    rq_activate_all_grippers(False)
    # end: URCap Program Node
  else:
    $ 55 "Else" "noBreak"
    # begin: URCap Program Node
    #   Source: Robotiq_Grippers, 3.17.0.105337, Robotiq Inc.
    #   Type: Gripper Activate
    $ 56 "Gripper Reset and Activate"

    kill rq_gripper_communication_thread
    rq_gripper_communication_thread_started = False
    rq_close_gripper_socket("1")
    rq_close_gripper_socket("2")
    rq_close_gripper_socket("3")
    rq_close_gripper_socket("4")

    rq_init_comm_if_connected(9, "1")
    rq_init_comm_if_connected(2, "2")
    rq_init_comm_if_connected(3, "3")
    rq_init_comm_if_connected(4, "4")
    rq_print_connected_grippers()
    rq_gripper_communication_thread = run rq_gripper_communication()

    while(not rq_gripper_communication_thread_started):
        sleep(0.008)
    end

    rq_set_max_current_for_all_grippers()

    reset_and_activate = True

    rq_activate_all_grippers(True)
    # end: URCap Program Node
  end
  $ 57 "zero_ftsensor()"
  zero_ftsensor()
  $ 58 "EXTT"
  $ 59 "Set GRP_3F_Enable=Off"
  set_standard_digital_out(4, False)
  $ 60 "Set BarcodeTrigger=Off"
  set_standard_digital_out(6, False)
  $ 61 "Set GRP_3F_Decap=Off"
  set_standard_digital_out(3, False)
  $ 62 "Set GRP_3F_Cap=Off"
  set_standard_digital_out(2, False)
  $ 63 "Set GRP_3F_Open=Off"
  set_standard_digital_out(5, False)
  $ 64 "PSE_T≔get_tool_free_pose(dir=[0,0,0.150], move_in_base_frame=True)"
  global PSE_T=get_tool_free_pose(dir=[0,0,0.150], move_in_base_frame=True)
  $ 65 "If is_reachable(Base_const, [PSE_T])"
  if (is_reachable(p[0.0,0.0,0.0,0.0,0.0,0.0], [PSE_T])):
    $ 66 "MoveL"
    $ 67 "PSE_T" "breakAfter"
    movel(PSE_T, a=1.2, v=0.15)
  end
  $ 68 "powder dispensing variable init"
  $ 69 "Start_thread≔ False "
  global Start_thread=  False
  $ 70 "vib_thread≔ False "
  global vib_thread=  False
  $ 71 "w_full_thread≔ False "
  global w_full_thread=  False
  $ 72 "d_cc≔0.07"
  global d_cc=0.07
  $ 73 "kp≔0.0035"
  global kp=0.0035
  $ 74 "ki≔0.0001"
  global ki=0.0001
  $ 75 "kd≔0.003"
  global kd=0.003
  $ 76 "dt≔0.2"
  global dt=0.2
  $ 77 "Integral_error≔0"
  global Integral_error=0
  $ 78 "current_error≔0"
  global current_error=0
  $ 79 "previous_error≔0"
  global previous_error=0
  $ 80 "tilt_increment≔0"
  global tilt_increment=0
  $ 81 "tilt_angle≔0"
  global tilt_angle=0
  $ 82 "diff≔0"
  global diff=0
  $ 83 "tilt_to_home()"
  tilt_to_home()
  $ 84 "tilt_to_home()"
  tilt_to_home()
  $ 85 "switch_spat_M≔ True "
  global switch_spat_M=  True
  $ 86 "switch_spat_S≔ True "
  global switch_spat_S=  True
  $ 87 "switch_spat_F_M≔ True "
  global switch_spat_F_M=  True
  $ 88 "switch_spat_F_S≔ True "
  global switch_spat_F_S=  True
  $ 89 "last_scale≔0"
  global last_scale=0
  $ 818 "Thread_1"
  thread Thread_1():
    while (True):
      $ 819 "Dosing Weight"
      $ 820 "If Start_thread≟ True "
      if (Start_thread ==   True  ):
        $ 821 "weight_value≔get_weight()"
        global weight_value=get_weight()
        $ 822 "diff≔target_weight-weight_value"
        global diff=target_weight-weight_value
        $ 823 "Wait: 0.2"
        sleep(0.2)
        $ 824 "sync()"
        sync()
      end
      $ 825 "sync()"
      sync()
    end
  end
  threadId_Thread_1 = run Thread_1()
  $ 826 "Thread_2"
  thread Thread_2():
    while (True):
      $ 827 "Vibration motor"
      $ 828 "Loop vib_thread≟ True "
      thread Thread_while_828():
        while (True):
          $ 829 "diff≔target_weight-weight_value"
          global diff=target_weight-weight_value
          $ 830 "If diff>0.02 and spatula≠'spatula_flat_S' "
          global thread_flag_830=0
          thread Thread_if_830():
            $ 832 "Set AO[0]=4.0"
            set_standard_analog_out(0, 0.4)
            thread_flag_830 = 1
          end
          if (diff>0.02  and  spatula != "spatula_flat_S" ):
            global thread_handler_830=run Thread_if_830()
            while (thread_flag_830 == 0):
              if not(diff>0.02  and  spatula != "spatula_flat_S" ):
                kill thread_handler_830
                thread_flag_830 = 2
              else:
                sync()
              end
            end
          else:
            thread_flag_830 = 2
          end
          if (thread_flag_830 == 2):
            $ 833 "ElseIf diff>0.02 and spatula≟'spatula_flat_S'"
            if (diff>0.02 and spatula == "spatula_flat_S"):
              $ 834 "vibration_3()"
              vibration_3()
            else:
              $ 835 "ElseIf diff≤0.03"
              global thread_flag_835=0
              thread Thread_if_835():
                $ 836 "vibration_2()"
                vibration_2()
                thread_flag_835 = 1
              end
              if (diff <= 0.03):
                global thread_handler_835=run Thread_if_835()
                while (thread_flag_835 == 0):
                  if not(diff <= 0.03):
                    kill thread_handler_835
                    thread_flag_835 = 2
                  else:
                    sync()
                  end
                end
              else:
                thread_flag_835 = 2
              end
              if (thread_flag_835 == 2):
                $ 837 "Else" "noBreak"
                $ 838 "Set AO[0]=0.0"
                set_standard_analog_out(0, 0.0)
              end
            end
          end
        end
      end
      if (vib_thread ==   True  ):
        global thread_handler_828=run Thread_while_828()
        while (vib_thread ==   True  ):
          sync()
        end
        kill thread_handler_828
      end
      $ 839 "sync()"
      sync()
    end
  end
  threadId_Thread_2 = run Thread_2()
  $ 840 "Thread_3"
  thread Thread_3():
    while (True):
      $ 841 "Container weight"
      $ 842 "If w_full_thread≟ True "
      if (w_full_thread ==   True  ):
        $ 843 "aa_weight_cont≔get_cont_weight()"
        global aa_weight_cont=get_cont_weight()
        $ 844 "Wait: 0.2"
        sleep(0.2)
        $ 845 "sync()"
        sync()
      end
      $ 846 "sync()"
      sync()
    end
  end
  threadId_Thread_3 = run Thread_3()
  while (True):
    $ 90 "Robot Program"
    $ 91 "MAIN"
    $ 92 "command_manager(external_control='uGO', cond_suspend=(ITM_Manipulated and AMR_AtTarget and AMR_Charging and AMR_Battery<40), cond_unsuspend=(AMR_Battery≟60))"
    command_manager(external_control="uGO", cond_suspend=(ITM_Manipulated  and  AMR_AtTarget  and  AMR_Charging  and  AMR_Battery<40), cond_unsuspend=(AMR_Battery == 60))
    $ 93 "log_state(STATE_Info)"
    log_state(STATE_Info)
    $ 94 "Switch STATE"
    switch_1 = STATE
    $ 95 "Case 1"
    if (1 == switch_1):
      $ 96 "Stopping"
      $ 97 "STATE_Info≔'Stopping'"
      global STATE_Info="Stopping"
      $ 98 "end_freedrive_mode()"
      end_freedrive_mode()
      $ 99 "Set"
      set_tcp(p[0.0,0.0,0.161,3.1415,0.0,0.0])
      $ 100 "PSE_T≔get_tool_free_pose(dir=[0,0,0.150], move_in_base_frame=True)"
      global PSE_T=get_tool_free_pose(dir=[0,0,0.150], move_in_base_frame=True)
      $ 101 "If is_reachable(Base_const, [PSE_T])"
      if (is_reachable(p[0.0,0.0,0.0,0.0,0.0,0.0], [PSE_T])):
        $ 102 "MoveL"
        $ 103 "PSE_T" "breakAfter"
        movel(PSE_T, a=1.2, v=0.15)
      end
      $ 104 "do_transition(keep_rxry=OBJ_Picked, r=0)"
      do_transition(keep_rxry=OBJ_Picked, r=0)
      $ 113 "Call Sub_AMR_MiR_V3"
      Sub_AMR_MiR_V3()
      $ 114 "If stopping() and AMR_Done"
      if (stopping()  and  AMR_Done):
        $ 115 "STATE≔2"
        global STATE=2
        $ 116 "ugo_update_outputs()"
        ugo_update_outputs()
      end
    elif (2 == switch_1):
      $ 117 "Case 2"
      $ 118 "Stopped"
      $ 119 "STATE_Info≔'Stopped'"
      global STATE_Info="Stopped"
      $ 120 "Call Sub_AMR_MiR_V3"
      Sub_AMR_MiR_V3()
      $ 121 "If CMD_Reset  or PB_Start"
      if (CMD_Reset   or  get_standard_digital_in(0)):
        $ 122 "STATE≔3"
        global STATE=3
        $ 123 "ugo_update_outputs()"
        ugo_update_outputs()
      end
    elif (3 == switch_1):
      $ 124 "Case 3"
      $ 125 " Resetting"
      $ 126 "STATE_Info≔'Resetting'"
      global STATE_Info="Resetting"
      $ 127 "uML"
      $ 128 "reset_error()"
      reset_error()
      $ 129 "reset_warning()"
      reset_warning()
      $ 130 "PROCESS_Step≔0"
      global PROCESS_Step=0
      $ 131 "PROCESS_Info≔''"
      global PROCESS_Info=""
      $ 132 "ARM_Referenced≔ False "
      global ARM_Referenced=  False
      $ 133 "WRK_Done≔ False "
      global WRK_Done=  False
      $ 134 "ITM_Prepared≔ False "
      global ITM_Prepared=  False
      $ 135 "ITM_Manipulated≔ False "
      global ITM_Manipulated=  False
      $ 136 "STP≔0"
      global STP=0
      $ 137 "Action≔0"
      global Action=0
      $ 138 "Action_Info≔''"
      global Action_Info=""
      $ 139 "ITM_ID≔0"
      global ITM_ID=0
      $ 140 "JIG≔0"
      global JIG=0
      $ 141 "JIG_Slot≔0"
      global JIG_Slot=0
      $ 142 "Task_info≔''"
      global Task_info=""
      $ 143 "Set"
      set_tcp(p[0.0,0.0,0.161,3.1415,0.0,0.0])
      $ 144 "App"
      $ 145 "'ADD APPLICATION SPECIFIC COMMANDS'"
      # 'ADD APPLICATION SPECIFIC COMMANDS'
      $ 146 "OBJ_Type≔0"
      global OBJ_Type=0
      $ 147 "OBJ_Nbr≔0"
      global OBJ_Nbr=0
      $ 148 "If CNT_Rack_Output≥50"
      if (CNT_Rack_Output >= 50):
        $ 149 "CNT_Rack_Output≔0"
        global CNT_Rack_Output=0
      end
      $ 150 "TASK≔struct(ID=0, NAVI=struct(target=0, footprint=0, protectiveOff=0, dock=0), WORK=struct(ITM_ID_Src=0, JIG_ID_Src=0, OBJ_Nbr_Src=0, ACT_Src=0, ITM_ID_Tgt=0, JIG_ID_Tgt=0, OBJ_Nbr_Tgt=0, ACT_Tgt=0, OBJ_Type=0))"
      global TASK=struct(ID=0, NAVI=struct(target=0, footprint=0, protectiveOff=0, dock=0), WORK=struct(ITM_ID_Src=0, JIG_ID_Src=0, OBJ_Nbr_Src=0, ACT_Src=0, ITM_ID_Tgt=0, JIG_ID_Tgt=0, OBJ_Nbr_Tgt=0, ACT_Tgt=0, OBJ_Type=0))
      $ 151 "Call Sub_AMR_MiR_V3"
      Sub_AMR_MiR_V3()
      $ 152 "If resetting() and AMR_Done"
      if (resetting()  and  AMR_Done):
        $ 153 "STATE≔4"
        global STATE=4
        $ 154 "ugo_update_outputs()"
        ugo_update_outputs()
      end
    elif (4 == switch_1):
      $ 155 "Case 4"
      $ 156 "Idle"
      $ 157 "STATE_Info≔'Idle'"
      global STATE_Info="Idle"
      $ 158 "If CMD_Start"
      if (CMD_Start):
        $ 159 "STATE≔5"
        global STATE=5
        $ 160 "ugo_update_outputs()"
        ugo_update_outputs()
      end
    elif (5 == switch_1):
      $ 161 "Case 5"
      $ 162 "Starting"
      $ 163 "STATE_Info≔'Starting'"
      global STATE_Info="Starting"
      $ 164 "'ADD COMMANDS WHAT TO START WITH'"
      # 'ADD COMMANDS WHAT TO START WITH'
      $ 165 "Call Sub_AMR_MiR_V3"
      Sub_AMR_MiR_V3()
      $ 166 "get ugo data"
      $ 167 "Assign Tasks"
      $ 168 "TASK.ID = ugo_get_task()"
      TASK.ID = ugo_get_task()
      $ 169 "If TASK.ID≟1"
      if (TASK.ID == 1):
        $ 170 "Task_info≔'Charge'"
        global Task_info="Charge"
        $ 171 "Parameters"
        $ 172 "AMR_PosTarget≔1"
        global AMR_PosTarget=1
      else:
        $ 173 "ElseIf TASK.ID≟9"
        if (TASK.ID == 9):
          $ 174 "'Pick Sarstedt Rack from Variable source'"
          # 'Pick Sarstedt Rack from Variable source'
          $ 175 "Task_info≔'Navigate to Target'"
          global Task_info="Navigate to Target"
          $ 176 "Parameters"
          $ 177 "AMR_PosTarget≔UGO.read_input('00','ITM_ID')"
          global AMR_PosTarget=UGO.read_input("00","ITM_ID")
        else:
          $ 178 "ElseIf TASK.ID≟13"
          if (TASK.ID == 13):
            $ 179 "Task_info≔'Dose Powder'"
            global Task_info="Dose Powder"
            $ 180 "Parameters"
            $ 181 "ITM_ID≔1"
            global ITM_ID=1
            $ 182 "W_now≔(UGO.read_input('00','Container_weight'))/1000"
            global W_now=(UGO.read_input("00","Container_weight"))/1000
            $ 183 "Pow_name≔(UGO.read_input('00','Powder_name'))"
            global Pow_name=(UGO.read_input("00","Powder_name"))
            $ 184 "target_weight≔(UGO.read_input('00','Target_weight'))/1000"
            global target_weight=(UGO.read_input("00","Target_weight"))/1000
            $ 185 "send_picking_info(Pow_name,target_weight)"
            send_picking_info(Pow_name,target_weight)
            $ 186 "w_dosed_total≔0"
            global w_dosed_total=0
            $ 187 "OBJ_Type≔6"
            global OBJ_Type=6
            $ 188 "JIG≔17"
            global JIG=17
            $ 189 "AMR_PosTarget≔5"
            global AMR_PosTarget=5
          else:
            $ 190 "ElseIf TASK.ID≟49"
            if (TASK.ID == 49):
              $ 191 "Task_info≔'Pick Containers'"
              global Task_info="Pick Containers"
              $ 192 "Parameters"
              $ 193 "ITM_ID≔1"
              global ITM_ID=1
              $ 194 "OBJ_Type≔6"
              global OBJ_Type=6
              $ 195 "JIG≔15"
              global JIG=15
              $ 196 "AMR_PosTarget≔3"
              global AMR_PosTarget=3
            else:
              $ 197 "ElseIf TASK.ID≟50"
              if (TASK.ID == 50):
                $ 198 "Task_info≔'Decap Containers'"
                global Task_info="Decap Containers"
                $ 199 "Parameters"
                $ 200 "ITM_ID≔1"
                global ITM_ID=1
                $ 201 "OBJ_Type≔6"
                global OBJ_Type=6
                $ 202 "JIG≔16"
                global JIG=16
                $ 203 "AMR_PosTarget≔5"
                global AMR_PosTarget=5
              else:
                $ 204 "ElseIf TASK.ID≟51"
                if (TASK.ID == 51):
                  $ 205 "Task_info≔'Detect Spatula and transfer powder'"
                  global Task_info="Detect Spatula and transfer powder"
                  $ 206 "Parameters"
                  $ 207 "ITM_ID≔1"
                  global ITM_ID=1
                  $ 208 "target_weight≔(UGO.read_input('00','Target_weight'))/1000"
                  global target_weight=(UGO.read_input("00","Target_weight"))/1000
                  $ 209 "OBJ_Type≔8"
                  global OBJ_Type=8
                  $ 210 "JIG≔16"
                  global JIG=16
                  $ 211 "AMR_PosTarget≔5"
                  global AMR_PosTarget=5
                else:
                  $ 212 "ElseIf TASK.ID≟52"
                  if (TASK.ID == 52):
                    $ 213 "Task_info≔'Pick Powder'"
                    global Task_info="Pick Powder"
                    $ 214 "Parameters"
                    $ 215 "ITM_ID≔1"
                    global ITM_ID=1
                    $ 217 "OBJ_Type≔6"
                    global OBJ_Type=6
                    $ 218 "JIG≔15"
                    global JIG=15
                    $ 219 "AMR_PosTarget≔3"
                    global AMR_PosTarget=3
                  else:
                    $ 220 "ElseIf TASK.ID≟53"
                    if (TASK.ID == 53):
                      $ 221 "Task_info≔'Decap Powder'"
                      global Task_info="Decap Powder"
                      $ 222 "Parameters"
                      $ 223 "ITM_ID≔1"
                      global ITM_ID=1
                      $ 224 "OBJ_Type≔6"
                      global OBJ_Type=6
                      $ 225 "JIG≔1"
                      global JIG=1
                      $ 226 "AMR_PosTarget≔5"
                      global AMR_PosTarget=5
                    else:
                      $ 227 "ElseIf TASK.ID≟54"
                      if (TASK.ID == 54):
                        $ 228 "Task_info≔'Empty and swap Powder container'"
                        global Task_info="Empty and swap Powder container"
                        $ 237 "Parameters"
                        $ 238 "ITM_ID≔1"
                        global ITM_ID=1
                        $ 240 "W_now≔(UGO.read_input('00','Container_weight'))/1000"
                        global W_now=(UGO.read_input("00","Container_weight"))/1000
                        $ 241 "Pow_name≔(UGO.read_input('00','Powder_name'))"
                        global Pow_name=(UGO.read_input("00","Powder_name"))
                        $ 244 "OBJ_Type≔6"
                        global OBJ_Type=6
                        $ 245 "JIG≔17"
                        global JIG=17
                        $ 246 "AMR_PosTarget≔5"
                        global AMR_PosTarget=5
                      else:
                        $ 247 "ElseIf TASK.ID≟55"
                        if (TASK.ID == 55):
                          $ 248 "Task_info≔'Place Powder'"
                          global Task_info="Place Powder"
                          $ 249 "Parameters"
                          $ 250 "ITM_ID≔1"
                          global ITM_ID=1
                          $ 251 "OBJ_Type≔6"
                          global OBJ_Type=6
                          $ 252 "JIG≔21"
                          global JIG=21
                          $ 253 "AMR_PosTarget≔5"
                          global AMR_PosTarget=5
                        else:
                          $ 254 "ElseIf TASK.ID≟56"
                          if (TASK.ID == 56):
                            $ 255 "Task_info≔'Dose Powder'"
                            global Task_info="Dose Powder"
                            $ 256 "Parameters"
                            $ 257 "ITM_ID≔1"
                            global ITM_ID=1
                            $ 258 "target_weight≔(UGO.read_input('00','Target_weight'))/1000"
                            global target_weight=(UGO.read_input("00","Target_weight"))/1000
                            $ 259 "W_now≔(UGO.read_input('00','Container_weight'))/1000"
                            global W_now=(UGO.read_input("00","Container_weight"))/1000
                            $ 260 "Pow_name≔(UGO.read_input('00','Powder_name'))"
                            global Pow_name=(UGO.read_input("00","Powder_name"))
                            $ 261 "OBJ_Type≔6"
                            global OBJ_Type=6
                            $ 262 "JIG≔17"
                            global JIG=17
                            $ 263 "AMR_PosTarget≔5"
                            global AMR_PosTarget=5
                          else:
                            $ 264 "ElseIf TASK.ID≟57"
                            if (TASK.ID == 57):
                              $ 265 "Task_info≔'Recipe Powder dosing'"
                              global Task_info="Recipe Powder dosing"
                              $ 266 "Parameters"
                              $ 267 "ITM_ID≔1"
                              global ITM_ID=1
                              $ 268 "Pow_A≔(UGO.read_input('00','PowderA'))"
                              global Pow_A=(UGO.read_input("00","PowderA"))
                              $ 269 "Pow_B≔(UGO.read_input('00','PowderB'))"
                              global Pow_B=(UGO.read_input("00","PowderB"))
                              $ 270 "Pow_C≔(UGO.read_input('00','PowderC'))"
                              global Pow_C=(UGO.read_input("00","PowderC"))
                              $ 271 "Total_weight≔(UGO.read_input('00','Total_weight'))/1000"
                              global Total_weight=(UGO.read_input("00","Total_weight"))/1000
                              $ 272 "Pow_A_percent≔(UGO.read_input('00','PowderA_percentage'))/100"
                              global Pow_A_percent=(UGO.read_input("00","PowderA_percentage"))/100
                              $ 273 "Pow_B_percent≔(UGO.read_input('00','PowderB_percentage'))/100"
                              global Pow_B_percent=(UGO.read_input("00","PowderB_percentage"))/100
                              $ 274 "Pow_C_percent≔(UGO.read_input('00','PowderC_percentage'))/100"
                              global Pow_C_percent=(UGO.read_input("00","PowderC_percentage"))/100
                              $ 275 "OBJ_Type≔6"
                              global OBJ_Type=6
                              $ 276 "JIG≔17"
                              global JIG=17
                              $ 277 "AMR_PosTarget≔5"
                              global AMR_PosTarget=5
                            else:
                              $ 278 "ElseIf TASK.ID≟58"
                              if (TASK.ID == 58):
                                $ 279 "Task_info≔'Pick Powder containers'"
                                global Task_info="Pick Powder containers"
                                $ 280 "Parameters"
                                $ 281 "ITM_ID≔1"
                                global ITM_ID=1
                                $ 282 "OBJ_Type≔6"
                                global OBJ_Type=6
                                $ 283 "JIG≔15"
                                global JIG=15
                                $ 284 "AMR_PosTarget≔3"
                                global AMR_PosTarget=3
                              else:
                                $ 285 "ElseIf TASK.ID≟59"
                                if (TASK.ID == 59):
                                  $ 286 "Task_info≔'Empty Powder container'"
                                  global Task_info="Empty Powder container"
                                  $ 287 "Parameters"
                                  $ 288 "ITM_ID≔1"
                                  global ITM_ID=1
                                  $ 290 "Pow_name≔(UGO.read_input('00','Powder_name'))"
                                  global Pow_name=(UGO.read_input("00","Powder_name"))
                                  $ 292 "target_weight≔aa_weight_cont-empty_weight_g"
                                  global target_weight=aa_weight_cont-empty_weight_g
                                  $ 293 "send_picking_info(Pow_name,target_weight)"
                                  send_picking_info(Pow_name,target_weight)
                                  $ 294 "w_dosed_total≔0"
                                  global w_dosed_total=0
                                  $ 295 "OBJ_Type≔6"
                                  global OBJ_Type=6
                                  $ 296 "JIG≔17"
                                  global JIG=17
                                  $ 297 "AMR_PosTarget≔5"
                                  global AMR_PosTarget=5
                                else:
                                  $ 298 "ElseIf TASK.ID≟61"
                                  if (TASK.ID == 61):
                                    $ 299 "Task_info≔'Weigh, Place & Decap'"
                                    global Task_info="Weigh, Place & Decap"
                                    $ 300 "Parameters"
                                    $ 301 "ITM_ID≔1"
                                    global ITM_ID=1
                                    $ 302 "OBJ_Type≔6"
                                    global OBJ_Type=6
                                    $ 303 "JIG≔21"
                                    global JIG=21
                                    $ 304 "AMR_PosTarget≔5"
                                    global AMR_PosTarget=5
                                  else:
                                    $ 305 "Else" "noBreak"
                                    $ 306 "set_error(ERROR_WRONG_ORDER)"
                                    set_error(ERROR_WRONG_ORDER)
                                  end
                                end
                              end
                            end
                          end
                        end
                      end
                    end
                  end
                end
              end
            end
          end
        end
      end
      $ 307 "test ugo"
      $ 308 "Wait: 0.2"
      sleep(0.2)
      $ 309 "ugo_update_outputs()"
      ugo_update_outputs()
      $ 310 "If starting() and AMR_Done"
      if (starting()  and  AMR_Done):
        $ 311 "log_message(Task_info, 'New Task: ')"
        log_message(Task_info, "New Task: ")
        $ 312 "log_message(to_str(TASK.ID), 'Task_ID: ')"
        log_message(to_str(TASK.ID), "Task_ID: ")
        $ 313 "do_transition(keep_rxry=OBJ_Picked)"
        do_transition(keep_rxry=OBJ_Picked)
        $ 314 "STATE≔6"
        global STATE=6
        $ 315 "ugo_update_outputs()"
        ugo_update_outputs()
      end
    elif (6 == switch_1):
      $ 316 "Case 6"
      $ 317 "Execute"
      $ 318 "STATE_Info≔'Execute'"
      global STATE_Info="Execute"
      $ 319 "If  not CMD_Hold and not CMD_Suspend"
      global thread_flag_319=0
      thread Thread_if_319():
        $ 320 "Switch PROCESS_Step"
        switch_2 = PROCESS_Step
        $ 321 "Case 0"
        if (0 == switch_2):
          $ 322 "PROCESS_Info≔'process control'"
          global PROCESS_Info="process control"
          $ 323 "log_process(PROCESS_Info)"
          log_process(PROCESS_Info)
          $ 324 "process control"
          $ 325 "If  not AMR_AtTarget"
          if (  not  AMR_AtTarget):
            $ 326 "PROCESS_Step≔1"
            global PROCESS_Step=1
          else:
            $ 327 "ElseIf (( not ITM_Prepared and  not WRK_Done) or (ITM_Prepared and WRK_Done))"
            if (((  not  ITM_Prepared  and    not  WRK_Done)  or  (ITM_Prepared  and  WRK_Done))):
              $ 328 "PROCESS_Step≔2"
              global PROCESS_Step=2
            else:
              $ 329 "ElseIf  not WRK_Done"
              if (  not  WRK_Done):
                $ 330 "PROCESS_Step≔3"
                global PROCESS_Step=3
              else:
                $ 331 "Else" "noBreak"
                $ 332 "task finished"
                $ 333 "PROCESS_Info≔''"
                global PROCESS_Info=""
                $ 334 "STATE≔7"
                global STATE=7
                $ 335 "ugo_update_outputs()"
                ugo_update_outputs()
              end
            end
          end
        elif (1 == switch_2):
          $ 336 "Case 1"
          $ 337 "navigate"
          $ 338 "'MOVING THE uML'"
          # 'MOVING THE uML'
          $ 339 "PROCESS_Info≔'move to target'"
          global PROCESS_Info="move to target"
          $ 340 "log_process(PROCESS_Info)"
          log_process(PROCESS_Info)
          $ 341 "If TASK.ID≟1"
          if (TASK.ID == 1):
            $ 342 "Action≔51"
            global Action=51
          else:
            $ 343 "Else" "noBreak"
            $ 344 "Action≔52"
            global Action=52
          end
          $ 345 "Call Sub_AMR_MiR_V3"
          Sub_AMR_MiR_V3()
          $ 346 "If AMR_Done"
          if (AMR_Done):
            $ 347 "PROCESS_Step≔0"
            global PROCESS_Step=0
          end
        elif (2 == switch_2):
          $ 348 "Case 2"
          $ 349 "prepare"
          $ 350 "'THINGS THAT HAVE TO BE DONE ONCE IN A SEQUENCE,WORKFLOW'"
          # 'THINGS THAT HAVE TO BE DONE ONCE IN A SEQUENCE,WORKFLOW'
          $ 351 "PROCESS_Info≔'prepare for work'"
          global PROCESS_Info="prepare for work"
          $ 352 "log_process(PROCESS_Info)"
          log_process(PROCESS_Info)
          $ 353 "If TASK.WORK.ITM_ID_Src>1"
          if (TASK.WORK.ITM_ID_Src>1):
            $ 354 "ITM_ID≔TASK.WORK.ITM_ID_Src"
            global ITM_ID=TASK.WORK.ITM_ID_Src
          else:
            $ 355 "ElseIf TASK.WORK.ITM_ID_Tgt>1"
            if (TASK.WORK.ITM_ID_Tgt>1):
              $ 356 "ITM_ID≔TASK.WORK.ITM_ID_Tgt"
              global ITM_ID=TASK.WORK.ITM_ID_Tgt
            end
          end
          $ 357 "If  not ARM_Referenced and (ITM_ID≠0)"
          if (  not  ARM_Referenced  and  (ITM_ID != 0)):
            $ 358 "STP≔1"
            global STP=1
          else:
            $ 359 "ElseIf ARM_Referenced or (ITM_ID≟0)"
            if (ARM_Referenced  or  (ITM_ID == 0)):
              $ 360 "STP≔2"
              global STP=2
            end
          end
          $ 361 "Switch STP"
          switch_3 = STP
          $ 362 "Case 1"
          if (1 == switch_3):
            $ 363 "reference"
            $ 364 "STP_Info≔'reference at target position'"
            global STP_Info="reference at target position"
            $ 365 "log_step(STP_Info)"
            log_step(STP_Info)
            $ 366 "If ITM_ID≟1"
            if (ITM_ID == 1):
              $ 367 "CAM_Done≔ True "
              global CAM_Done=  True
            else:
              $ 368 "Else" "noBreak"
              $ 369 "Action≔131"
              global Action=131
              $ 370 "Call Sub_Vision_V18"
              Sub_Vision_V18()
            end
            $ 372 "If CAM_Done and  not ERROR.FLAG"
            if (CAM_Done  and    not  ERROR.FLAG):
              $ 373 "log_step('ARM referenced')"
              log_step("ARM referenced")
              $ 374 "ARM_Referenced≔ True "
              global ARM_Referenced=  True
            end
          elif (2 == switch_3):
            $ 375 "Case 2"
            $ 376 "manipulate"
            $ 377 "STP_Info≔'manipulate item'"
            global STP_Info="manipulate item"
            $ 378 "log_step(STP_Info)"
            log_step(STP_Info)
            $ 379 "'In case pressing button is needed'"
            # 'In case pressing button is needed'
            $ 380 "If found_in_list(ITM_ID, ITM_ID_List)"
            if (found_in_list(ITM_ID, ITM_ID_List)):
              $ 381 "Switch ITM_ID"
              switch_4 = ITM_ID
              $ 382 "Case 0"
              if (0 == switch_4):
                $ 383 "ITM_Manipulated≔ not ITM_Manipulated"
                global ITM_Manipulated=  not  ITM_Manipulated
              elif (1 == switch_4):
                $ 384 "Case 1"
                $ 385 "ITM_Manipulated≔ not ITM_Manipulated"
                global ITM_Manipulated=  not  ITM_Manipulated
              elif (2 == switch_4):
                $ 386 "Case 2"
              else:
                $ 396 "Default Case"
                $ 397 "ITM_Manipulated≔ not ITM_Manipulated"
                global ITM_Manipulated=  not  ITM_Manipulated
              end
            end
          end
          $ 398 "ITM_Prepared≔(ITM_Manipulated or  not found_in_list(ITM_ID, ITM_ID_List)) and (ARM_Referenced or ITM_ID≟0) and  not WRK_Done"
          global ITM_Prepared=(ITM_Manipulated  or    not  found_in_list(ITM_ID, ITM_ID_List))  and  (ARM_Referenced  or  ITM_ID == 0)  and    not  WRK_Done
          $ 399 "STP≔0"
          global STP=0
          $ 400 "STP_Info≔''"
          global STP_Info=""
          $ 401 "PROCESS_Step≔0"
          global PROCESS_Step=0
        elif (3 == switch_2):
          $ 402 "Case 3"
          $ 403 "work"
          $ 404 "'ADD EVERY MACHINE, OBJECT, STATION TO WORK ON'"
          # 'ADD EVERY MACHINE, OBJECT, STATION TO WORK ON'
          $ 405 "Switch ITM_ID"
          switch_3 = ITM_ID
          $ 406 "Case 1"
          if (1 == switch_3):
            $ 407 "uLM"
            $ 408 "If TASK.ID≟12"
            if (TASK.ID == 12):
              $ 409 "fill racks"
              $ 410 "Action≔151"
              global Action=151
              $ 411 "Call Sub_Vision_V18"
              Sub_Vision_V18()
              $ 412 "If  not ERROR.FLAG"
              if (  not  ERROR.FLAG):
                $ 413 "Actions for the task"
                $ 414 "Action≔1"
                global Action=1
                $ 415 "JIG≔2"
                global JIG=2
                $ 416 "JIG_Slot≔CAM_Result[0]"
                global JIG_Slot=CAM_Result[0]
                $ 417 "OBJ_Nbr≔CAM_Result[0]"
                global OBJ_Nbr=CAM_Result[0]
                $ 418 "OBJ_Type≔2"
                global OBJ_Type=2
                $ 419 "Call Sub_Action_V4"
                Sub_Action_V4()
                $ 420 "If OBJ_Picked"
                if (OBJ_Picked):
                  $ 421 "CAM_Result.remove(0)"
                  CAM_Result.remove(0)
                  $ 422 "PRC_TubCounter≔PRC_TubCounter+1"
                  global PRC_TubCounter=PRC_TubCounter+1
                  $ 423 "If PRC_TubCounter%4≟0"
                  if (PRC_TubCounter%4 == 0):
                    $ 424 "JIG_Slot≔4"
                    global JIG_Slot=4
                  else:
                    $ 425 "Else" "noBreak"
                    $ 426 "JIG_Slot≔PRC_TubCounter%4"
                    global JIG_Slot=PRC_TubCounter%4
                  end
                  $ 427 "OBJ_Nbr≔ceil(PRC_TubCounter/4)"
                  global OBJ_Nbr=ceil(PRC_TubCounter/4)
                  $ 428 "Action≔2"
                  global Action=2
                  $ 429 "JIG≔4"
                  global JIG=4
                  $ 430 "Call Sub_Action_V4"
                  Sub_Action_V4()
                  $ 431 "Action≔151"
                  global Action=151
                  $ 432 "Call Sub_Vision_V18"
                  Sub_Vision_V18()
                end
              end
              $ 433 "If (CAM_Captures≥CAM_PRM_Retries) or (PRC_TubCounter≥32)"
              if ((CAM_Captures >= CAM_PRM_Retries)  or  (PRC_TubCounter >= 32)):
                $ 434 "PROCESS_Step≔0"
                global PROCESS_Step=0
                $ 435 "WRK_Done≔ True "
                global WRK_Done=  True
              end
            else:
              $ 436 "ElseIf TASK.ID≟13"
              if (TASK.ID == 13):
                $ 437 "Dose Powder"
                $ 438 "Action≔131"
                global Action=131
                $ 439 "Call Sub_Vision_V18"
                Sub_Vision_V18()
                $ 440 "Action≔34"
                global Action=34
                $ 441 "Call Sub_Action_V4"
                Sub_Action_V4()
                $ 442 "PROCESS_Step≔0"
                global PROCESS_Step=0
                $ 443 "WRK_Done≔ True "
                global WRK_Done=  True
              else:
                $ 444 "ElseIf TASK.ID≟49"
                if (TASK.ID == 49):
                  $ 445 "Pick Powder container"
                  $ 446 "Action≔131"
                  global Action=131
                  $ 447 "Call Sub_Vision_V18"
                  Sub_Vision_V18()
                  $ 448 "Action≔35"
                  global Action=35
                  $ 449 "Call Sub_Action_V4"
                  Sub_Action_V4()
                  $ 450 "PROCESS_Step≔0"
                  global PROCESS_Step=0
                  $ 451 "WRK_Done≔ True "
                  global WRK_Done=  True
                else:
                  $ 452 "ElseIf TASK.ID≟50"
                  if (TASK.ID == 50):
                    $ 453 "Decap containers"
                    $ 454 "Action≔36"
                    global Action=36
                    $ 455 "Call Sub_Action_V4"
                    Sub_Action_V4()
                    $ 456 "PROCESS_Step≔0"
                    global PROCESS_Step=0
                    $ 457 "WRK_Done≔ True "
                    global WRK_Done=  True
                  else:
                    $ 458 "ElseIf TASK.ID≟51"
                    if (TASK.ID == 51):
                      $ 459 "Detect Spatula and transfer powder"
                      $ 460 "Action≔131"
                      global Action=131
                      $ 461 "Call Sub_Vision_V18"
                      Sub_Vision_V18()
                      $ 462 "Action≔37"
                      global Action=37
                      $ 463 "Call Sub_Action_V4"
                      Sub_Action_V4()
                      $ 464 "PROCESS_Step≔0"
                      global PROCESS_Step=0
                      $ 465 "WRK_Done≔ True "
                      global WRK_Done=  True
                    else:
                      $ 466 "ElseIf TASK.ID≟52"
                      if (TASK.ID == 52):
                        $ 467 "Pick Powder container"
                        $ 468 "Action≔131"
                        global Action=131
                        $ 469 "Call Sub_Vision_V18"
                        Sub_Vision_V18()
                        $ 470 "Action≔39"
                        global Action=39
                        $ 471 "Call Sub_Action_V4"
                        Sub_Action_V4()
                        $ 472 "PROCESS_Step≔0"
                        global PROCESS_Step=0
                        $ 473 "WRK_Done≔ True "
                        global WRK_Done=  True
                      else:
                        $ 474 "ElseIf TASK.ID≟53"
                        if (TASK.ID == 53):
                          $ 475 "Decap containerA"
                          $ 476 "Action≔40"
                          global Action=40
                          $ 477 "Call Sub_Action_V4"
                          Sub_Action_V4()
                          $ 478 "PROCESS_Step≔0"
                          global PROCESS_Step=0
                          $ 479 "WRK_Done≔ True "
                          global WRK_Done=  True
                        else:
                          $ 480 "ElseIf TASK.ID≟55"
                          if (TASK.ID == 55):
                            $ 481 "Place Powder"
                            $ 482 "Action≔131"
                            global Action=131
                            $ 483 "Call Sub_Vision_V18"
                            Sub_Vision_V18()
                            $ 484 "Action≔41"
                            global Action=41
                            $ 485 "Call Sub_Action_V4"
                            Sub_Action_V4()
                            $ 486 "PROCESS_Step≔0"
                            global PROCESS_Step=0
                            $ 487 "WRK_Done≔ True "
                            global WRK_Done=  True
                          else:
                            $ 488 "ElseIf TASK.ID≟54"
                            if (TASK.ID == 54):
                              $ 489 "Empty and swap container"
                              $ 490 "Action≔131"
                              global Action=131
                              $ 491 "Call Sub_Vision_V18"
                              Sub_Vision_V18()
                              $ 492 "Action≔42"
                              global Action=42
                              $ 493 "Call Sub_Action_V4"
                              Sub_Action_V4()
                              $ 494 "PROCESS_Step≔0"
                              global PROCESS_Step=0
                              $ 495 "WRK_Done≔ True "
                              global WRK_Done=  True
                            else:
                              $ 496 "ElseIf TASK.ID≟56"
                              if (TASK.ID == 56):
                                $ 497 "Dispense Powder"
                                $ 498 "Action≔131"
                                global Action=131
                                $ 499 "Call Sub_Vision_V18"
                                Sub_Vision_V18()
                                $ 500 "Action≔43"
                                global Action=43
                                $ 501 "Call Sub_Action_V4"
                                Sub_Action_V4()
                                $ 502 "PROCESS_Step≔0"
                                global PROCESS_Step=0
                                $ 503 "WRK_Done≔ True "
                                global WRK_Done=  True
                              else:
                                $ 504 "ElseIf TASK.ID≟57"
                                if (TASK.ID == 57):
                                  $ 505 "Recipe Dosing"
                                  $ 506 "Action≔48"
                                  global Action=48
                                  $ 507 "Call Sub_Action_V4"
                                  Sub_Action_V4()
                                  $ 524 "PROCESS_Step≔0"
                                  global PROCESS_Step=0
                                  $ 525 "WRK_Done≔ True "
                                  global WRK_Done=  True
                                else:
                                  $ 526 "ElseIf TASK.ID≟58"
                                  if (TASK.ID == 58):
                                    $ 527 "Pick Powder containers"
                                    $ 528 "Num_cont_picked≔0"
                                    global Num_cont_picked=0
                                    $ 529 "powder_position≔'Position1'"
                                    global powder_position="Position1"
                                    $ 530 "Loop Num_cont_picked<3"
                                    while (Num_cont_picked<3):
                                      $ 531 "Action≔131"
                                      global Action=131
                                      $ 532 "Call Sub_Vision_V18"
                                      Sub_Vision_V18()
                                      $ 533 "Action≔47"
                                      global Action=47
                                      $ 534 "Call Sub_Action_V4"
                                      Sub_Action_V4()
                                    end
                                    $ 535 "PROCESS_Step≔0"
                                    global PROCESS_Step=0
                                    $ 536 "WRK_Done≔ True "
                                    global WRK_Done=  True
                                  else:
                                    $ 537 "ElseIf TASK.ID≟59"
                                    if (TASK.ID == 59):
                                      $ 538 "Empty powder container"
                                      $ 539 "Action≔131"
                                      global Action=131
                                      $ 540 "Call Sub_Vision_V18"
                                      Sub_Vision_V18()
                                      $ 541 "Action≔50"
                                      global Action=50
                                      $ 542 "Call Sub_Action_V4"
                                      Sub_Action_V4()
                                      $ 543 "PROCESS_Step≔0"
                                      global PROCESS_Step=0
                                      $ 544 "WRK_Done≔ True "
                                      global WRK_Done=  True
                                    else:
                                      $ 545 "ElseIf TASK.ID≟61"
                                      if (TASK.ID == 61):
                                        $ 546 "Place Powder"
                                        $ 547 "Action≔131"
                                        global Action=131
                                        $ 548 "Call Sub_Vision_V18"
                                        Sub_Vision_V18()
                                        $ 549 "Action≔51"
                                        global Action=51
                                        $ 550 "Call Sub_Action_V4"
                                        Sub_Action_V4()
                                        $ 551 "PROCESS_Step≔0"
                                        global PROCESS_Step=0
                                        $ 552 "WRK_Done≔ True "
                                        global WRK_Done=  True
                                      end
                                    end
                                  end
                                end
                              end
                            end
                          end
                        end
                      end
                    end
                  end
                end
              end
            end
          elif (2 == switch_3):
            $ 553 "Case 2"
          elif (5 == switch_3):
            $ 595 "Case 5"
          elif (20 == switch_3):
            $ 603 "Case 20"
          elif (43 == switch_3):
            $ 665 "Case 43"
          else:
            $ 673 "Default Case"
            $ 674 "WRK_Done≔ True "
            global WRK_Done=  True
            $ 675 "PROCESS_Step≔0"
            global PROCESS_Step=0
          end
        end
        thread_flag_319 = 1
      end
      if (  not  CMD_Hold and not CMD_Suspend):
        global thread_handler_319=run Thread_if_319()
        while (thread_flag_319 == 0):
          if not(  not  CMD_Hold and not CMD_Suspend):
            kill thread_handler_319
            thread_flag_319 = 2
          else:
            sync()
          end
        end
      else:
        thread_flag_319 = 2
      end
      $ 676 "If CMD_Hold"
      if (CMD_Hold):
        $ 677 "STATE≔9"
        global STATE=9
        $ 678 "ugo_update_outputs()"
        ugo_update_outputs()
      else:
        $ 679 "ElseIf CMD_Suspend"
        if (CMD_Suspend):
          $ 680 "STATE≔12"
          global STATE=12
          $ 681 "ugo_update_outputs()"
          ugo_update_outputs()
        end
      end
    elif (7 == switch_1):
      $ 682 "Case 7"
      $ 683 "Completing"
      $ 684 "STATE_Info≔'Completing'"
      global STATE_Info="Completing"
      $ 685 "'ADD COMMANDS FOR COMPLETING THE PROCESS'"
      # 'ADD COMMANDS FOR COMPLETING THE PROCESS'
      $ 686 "do_transition(keep_rxry=OBJ_Picked)"
      do_transition(keep_rxry=OBJ_Picked)
      $ 687 "Call Sub_AMR_MiR_V3"
      Sub_AMR_MiR_V3()
      $ 688 "If completing() and AMR_Done"
      if (completing()  and  AMR_Done):
        $ 689 "STATE≔8"
        global STATE=8
        $ 690 "ugo_update_outputs()"
        ugo_update_outputs()
      end
    elif (8 == switch_1):
      $ 691 "Case 8"
      $ 692 "Complete"
      $ 693 "STATE_Info≔'Complete'"
      global STATE_Info="Complete"
      $ 694 "If CMD_Reset"
      if (CMD_Reset):
        $ 695 "STATE≔3"
        global STATE=3
        $ 696 "ugo_update_outputs()"
        ugo_update_outputs()
      end
    elif (9 == switch_1):
      $ 697 "Case 9"
      $ 698 "Holding"
      $ 699 "STATE_Info≔'Holding'"
      global STATE_Info="Holding"
      $ 700 "stopl(0.5)"
      stopl(0.5)
      $ 701 "Call Sub_AMR_MiR_V3"
      Sub_AMR_MiR_V3()
      $ 702 "If holding() and AMR_Done"
      if (holding()  and  AMR_Done):
        $ 703 "STATE≔10"
        global STATE=10
        $ 704 "ugo_update_outputs()"
        ugo_update_outputs()
      end
    elif (10 == switch_1):
      $ 705 "Case 10"
      $ 706 "Held"
      $ 707 "STATE_Info≔'Held'"
      global STATE_Info="Held"
      $ 708 "If CMD_Unhold"
      if (CMD_Unhold):
        $ 709 "end_freedrive_mode()"
        end_freedrive_mode()
        $ 710 "STATE≔11"
        global STATE=11
        $ 711 "ugo_update_outputs()"
        ugo_update_outputs()
      else:
        $ 712 "ElseIf FNC_Freedrive"
        if (FNC_Freedrive):
          $ 713 "freedrive_mode()"
          freedrive_mode()
        else:
          $ 714 "Else" "noBreak"
          $ 715 "end_freedrive_mode()"
          end_freedrive_mode()
        end
      end
    elif (11 == switch_1):
      $ 716 "Case 11"
      $ 717 "Unholding"
      $ 718 "STATE_Info≔'Unholding'"
      global STATE_Info="Unholding"
      $ 719 "Clearing"
      $ 720 "Switch ERROR.ID"
      switch_2 = ERROR.ID
      $ 721 "Case 1002"
      if (1002 == switch_2):
        $ 722 "AMR_AtTarget≔ False "
        global AMR_AtTarget=  False
        $ 723 "ARM_Referenced≔ False "
        global ARM_Referenced=  False
        $ 724 "ITM_Prepared≔ False "
        global ITM_Prepared=  False
        $ 725 "PROCESS_Step≔1"
        global PROCESS_Step=1
      elif (2007 == switch_2):
        $ 726 "Case 2007"
        $ 727 "PROCESS_Step≔1"
        global PROCESS_Step=1
      end
      $ 728 "reset_error()"
      reset_error()
      $ 729 "reset_warning()"
      reset_warning()
      $ 730 "OBJ_Picked≔gripper_has_object()"
      global OBJ_Picked=gripper_has_object()
      $ 731 "Call Sub_AMR_MiR_V3"
      Sub_AMR_MiR_V3()
      $ 732 "If unholding() and AMR_Done"
      if (unholding()  and  AMR_Done):
        $ 733 "STATE≔6"
        global STATE=6
        $ 734 "ugo_update_outputs()"
        ugo_update_outputs()
      end
    elif (12 == switch_1):
      $ 735 "Case 12"
      $ 736 "Suspending"
      $ 737 "STATE_Info≔'Suspending'"
      global STATE_Info="Suspending"
      $ 738 "PROCESS_Info≔str_cat(PROCESS_Info, ' suspended')"
      global PROCESS_Info=str_cat(PROCESS_Info, " suspended")
      $ 739 "If suspending()"
      if (suspending()):
        $ 740 "STATE≔13"
        global STATE=13
        $ 741 "ugo_update_outputs()"
        ugo_update_outputs()
      end
    elif (13 == switch_1):
      $ 742 "Case 13"
      $ 743 "Suspended"
      $ 744 "STATE_Info≔'Suspended'"
      global STATE_Info="Suspended"
      $ 745 "Call Sub_AMR_MiR_V3"
      Sub_AMR_MiR_V3()
      $ 746 "If CMD_Unsuspend"
      if (CMD_Unsuspend):
        $ 747 "STATE≔14"
        global STATE=14
        $ 748 "ugo_update_outputs()"
        ugo_update_outputs()
      end
    elif (14 == switch_1):
      $ 749 "Case 14"
      $ 750 "Unsuspending"
      $ 751 "STATE_Info≔'Unsuspending'"
      global STATE_Info="Unsuspending"
      $ 752 "PROCESS_Step≔0"
      global PROCESS_Step=0
      $ 753 "If unsuspending()"
      if (unsuspending()):
        $ 754 "STATE≔6"
        global STATE=6
        $ 755 "ugo_update_outputs()"
        ugo_update_outputs()
      end
    elif (15 == switch_1):
      $ 756 "Case 15"
      $ 757 "Aborting"
      $ 758 "STATE_Info≔'Aborting'"
      global STATE_Info="Aborting"
      $ 759 "If aborting()"
      if (aborting()):
        $ 760 "STATE≔16"
        global STATE=16
        $ 761 "ugo_update_outputs()"
        ugo_update_outputs()
      end
    elif (16 == switch_1):
      $ 762 "Case 16"
      $ 763 "Aborted"
      $ 764 "STATE_Info≔'Aborted'"
      global STATE_Info="Aborted"
      $ 765 "If CMD_Clear"
      if (CMD_Clear):
        $ 766 "STATE≔17"
        global STATE=17
        $ 767 "ugo_update_outputs()"
        ugo_update_outputs()
      end
    elif (17 == switch_1):
      $ 768 "Case 17"
      $ 769 "Clearing"
      $ 770 "STATE_Info≔'Clearing'"
      global STATE_Info="Clearing"
      $ 771 "Clearing"
      $ 772 "reset_warning()"
      reset_warning()
      $ 773 "reset_error()"
      reset_error()
      $ 774 "If clearing()"
      if (clearing()):
        $ 775 "STATE≔2"
        global STATE=2
        $ 776 "ugo_update_outputs()"
        ugo_update_outputs()
      end
    end
    $ 777 "log_state(STATE_Info)"
    log_state(STATE_Info)
    $ 778 "log_warning(WARNING.MSG)"
    log_warning(WARNING.MSG)
    $ 779 "log_error(ERROR.MSG)"
    log_error(ERROR.MSG)
    $ 780 "Times"
    $ 781 "Switch STATE"
    switch_1 = STATE
    $ 782 "Case 1"
    if (1 == switch_1):
      $ 783 "TM_St_Stopping≔get_time(STATE_Times[STATE-1])"
      global TM_St_Stopping=get_time(STATE_Times[STATE-1])
    elif (2 == switch_1):
      $ 784 "Case 2"
      $ 785 "TM_St_Stopped≔get_time(STATE_Times[STATE-1])"
      global TM_St_Stopped=get_time(STATE_Times[STATE-1])
    elif (3 == switch_1):
      $ 786 "Case 3"
      $ 787 "TM_St_Resetting≔get_time(STATE_Times[STATE-1])"
      global TM_St_Resetting=get_time(STATE_Times[STATE-1])
    elif (4 == switch_1):
      $ 788 "Case 4"
      $ 789 "TM_St_Idle≔get_time(STATE_Times[STATE-1])"
      global TM_St_Idle=get_time(STATE_Times[STATE-1])
    elif (5 == switch_1):
      $ 790 "Case 5"
      $ 791 "TM_St_Starting≔get_time(STATE_Times[STATE-1])"
      global TM_St_Starting=get_time(STATE_Times[STATE-1])
    elif (6 == switch_1):
      $ 792 "Case 6"
      $ 793 "TM_St_Execute≔get_time(STATE_Times[STATE-1])"
      global TM_St_Execute=get_time(STATE_Times[STATE-1])
    elif (7 == switch_1):
      $ 794 "Case 7"
      $ 795 "TM_St_Completin≔get_time(STATE_Times[STATE-1])"
      global TM_St_Completin=get_time(STATE_Times[STATE-1])
    elif (8 == switch_1):
      $ 796 "Case 8"
      $ 797 "TM_St_Complete≔get_time(STATE_Times[STATE-1])"
      global TM_St_Complete=get_time(STATE_Times[STATE-1])
    elif (9 == switch_1):
      $ 798 "Case 9"
      $ 799 "TM_St_Holding≔get_time(STATE_Times[STATE-1])"
      global TM_St_Holding=get_time(STATE_Times[STATE-1])
    elif (10 == switch_1):
      $ 800 "Case 10"
      $ 801 "TM_St_Held≔get_time(STATE_Times[STATE-1])"
      global TM_St_Held=get_time(STATE_Times[STATE-1])
    elif (11 == switch_1):
      $ 802 "Case 11"
      $ 803 "TM_St_Unholding≔get_time(STATE_Times[STATE-1])"
      global TM_St_Unholding=get_time(STATE_Times[STATE-1])
    elif (12 == switch_1):
      $ 804 "Case 12"
      $ 805 "TM_St_Suspendin≔get_time(STATE_Times[STATE-1])"
      global TM_St_Suspendin=get_time(STATE_Times[STATE-1])
    elif (13 == switch_1):
      $ 806 "Case 13"
      $ 807 "TM_St_Suspended≔get_time(STATE_Times[STATE-1])"
      global TM_St_Suspended=get_time(STATE_Times[STATE-1])
    elif (14 == switch_1):
      $ 808 "Case 14"
      $ 809 "TM_St_Unsuspend≔get_time(STATE_Times[STATE-1])"
      global TM_St_Unsuspend=get_time(STATE_Times[STATE-1])
    elif (15 == switch_1):
      $ 810 "Case 15"
      $ 811 "TM_St_Aborting≔get_time(STATE_Times[STATE-1])"
      global TM_St_Aborting=get_time(STATE_Times[STATE-1])
    elif (16 == switch_1):
      $ 812 "Case 16"
      $ 813 "TM_St_Aborted≔get_time(STATE_Times[STATE-1])"
      global TM_St_Aborted=get_time(STATE_Times[STATE-1])
    elif (17 == switch_1):
      $ 814 "Case 17"
      $ 815 "TM_St_Clearing≔get_time(STATE_Times[STATE-1])"
      global TM_St_Clearing=get_time(STATE_Times[STATE-1])
    end
    $ 817 "Wait: 0.1"
    sleep(0.1)
  end
end
